FUNCTION_BLOCK FB_CoverClosingState EXTENDS FB_CoverState
VAR
	nStage			: UINT:= 0;
	tonDelta		: TON;		// PT is taken from pCover^.Delta at the start of each cycle (#76)
	tonFullCycle	: TON;		// PT is taken from pCover^.TimeToCycle at the start of each cycle (#76)
END_VAR

METHOD OpenCommand : BOOL
nStage := 0;
tonDelta(IN:=FALSE);
tonFullCycle(IN:=FALSE);
pCover^.SetState(pCover^.fbCoverOpeningState);
END_METHOD

METHOD RunState : BOOL
tonDelta();
tonFullCycle();
CASE nStage OF
	0:
		// #76: the cycle times were only read once, by the declaration initialisers, so the inputs of FB_CoverControl
		// never reached the timers. Take them at the start of each cycle (not every scan: a change mid-cycle must not
		// end it early).
		tonDelta.PT := pCover^.Delta;
		IF pCover^.TimeToCycle > T#0S THEN
			tonFullCycle.PT := pCover^.TimeToCycle;
		ELSE
			tonFullCycle.PT := T#15S;	// 0 would declare the end position after one scan
		END_IF
		pCover^._CoverState := E_MirrorCoverState.closing;
		tonDelta.IN := TRUE;
		nStage := 1;
	1:
		// Stop Motor 1
		pCover^._Motor1RelaisA := FALSE;
		pCover^._Motor1RelaisB := FALSE;
		// Close Motor 2
		pCover^._Motor2RelaisA := FALSE;
		pCover^._Motor2RelaisB := TRUE;
		nStage := 2;
	2:
		IF tonDelta.Q THEN
			tonDelta.IN := FALSE;
			nStage:=3;
		END_IF 
	3:
		// Close Motor 1
		pCover^._Motor1RelaisA := FALSE;
		pCover^._Motor1RelaisB := TRUE;
		tonFullCycle.IN:=TRUE;
		nStage := 4;
	4:
		IF tonFullCycle.Q THEN
			tonFullCycle.IN := FALSE;
			THIS^.SuccessfulFinished();
		END_IF 
END_CASE
END_METHOD

METHOD StopCommand : BOOL
nStage := 0;
tonDelta(IN:=FALSE);
tonFullCycle(IN:=FALSE);
pCover^.SetState(pCover^.fbCoverStoppingState);
END_METHOD

METHOD SuccessfulFinished : BOOL
nStage := 0;
tonDelta(IN:=FALSE);
tonFullCycle(IN:=FALSE);
// #71: release the relays at the end position (limit switches cut the motors, the covers are self-locking)
pCover^._Motor1RelaisA := FALSE;
pCover^._Motor1RelaisB := FALSE;
pCover^._Motor2RelaisA := FALSE;
pCover^._Motor2RelaisB := FALSE;
pCover^._CoverState := E_MirrorCoverState.closed;
pCover^.SetState(pCover^.fbCoverIdleState);
END_METHOD

END_FUNCTION_BLOCK

(* stored: Version 1.1.0.1, ProductVersion 3.1.4024.15
   POU FB_CoverClosingState: Id {01dc9b33-581a-47c6-88d3-673a749ad1ec}, SpecialFunc None
   Method OpenCommand: Id {37b09ab2-b8c8-4a93-a138-b28f6cb2bcf3}
   Method RunState: Id {80955472-6560-4181-a9ba-febd31ed8ad0}
   Method StopCommand: Id {81fd907d-7afe-4d61-9013-3ad196b8d9b7}
   Method SuccessfulFinished: Id {9a7dbaad-c9df-40cc-bdd5-9cc345f04d2e} *)
